VAR_GLOBAL
    bLowerButton : BOOL;
    bUpperButton : BOOL;
    bLightRelay : BOOL;
    bTemporaryLightRelay : BOOL;
END_VAR

(* stored: Version 1.1.0.1
   GVL GVL_EntrywaySimulation: Id {72DAEA00-AA6D-4DC6-904D-FDBF7FF27CBA} *)
